(* CODESYS project P_InstanceName.xml

Project tree, tasks and I/O mapping:
*)

// P_InstanceName
PROPERTY P_InstanceName : STRING
END_PROPERTY
